// TIA Portal V20 export
// export: Created 2026-10-20T12:52:58.7186213Z, ExportSetting WithDefaults, DisplayName Totally Integrated Automation Portal, DisplayVersion V20 Update 6, DisplayName TIA Portal Openness, DisplayVersion V20 Update 6, DisplayName TIA Portal Version Control Interface, DisplayVersion V20 Update 6, DisplayName SINAMICS Startdrive Advanced, DisplayVersion V20 SP1, DisplayName SINAMICS Startdrive G130, G150, S120, S150, SINAMICS MV, G220, S200, S210, DisplayVersion V20 SP1, DisplayName SINAMICS Startdrive G110M, G120, G120C, G120D, G120P, G115D, DisplayVersion V20 SP1, DisplayName STEP 7 Professional, DisplayVersion V20 Update 6, DisplayName STEP 7 Safety, DisplayVersion V20 Update 2, DisplayName WinCC Basic/Comfort/Advanced, DisplayVersion V20 Update 6, DisplayName WinCC Unified, DisplayVersion V20 Update 6
DATA_BLOCK "DB_Send_Data_To_Logistex"   // DB901
{ S7_Optimized_Access := 'TRUE' }
VERSION : 0.1
// stored: AutoNumber false, DBAccessibleFromOPCUA true, IsOnlyStoredInLoadMemory false, IsRetainMemResEnabled false, IsWriteProtectedInAS false, MemoryReserve 100
   VAR
      VTD_J1310_INFEED : "VTD_Infeed";
      VTD_J1320_INFEED { S7_SetPoint := 'True'} : "VTD_Infeed";
      VTD_J1330_INFEED { S7_SetPoint := 'True'} : "VTD_Infeed";
      VTD_J1310_OUTFEED { S7_SetPoint := 'True'} : "VTD_Outfeed";
      VTD_J1320_OUTFEED { S7_SetPoint := 'True'} : "VTD_Outfeed";
      VTD_J1330_OUTFEED { S7_SetPoint := 'True'} : "VTD_Outfeed";
      VTD_STATUS : Array[1..10] of Byte;
      PLC_STATUS : Struct
         Hardbit : Bool;
         "PLC_E-Stop" : Bool;
      END_STRUCT;
      CONV_SPEED : Struct
         VTD_J1310_INF_SP : Int;
         VTD_J1310_OUF_SP : Int;
         VTD_J1320_INF_SP : Int;
         VTD_J1320_OUF_SP : Int;
         VTD_J1330_INF_SP_1 : Int;
         VTD_J1330_OUF_SP : Int;
      END_STRUCT;
   END_VAR
BEGIN
END_DATA_BLOCK
